(* IEC 61131-3 sources: Lasal-MCP/examples/SampleSource/LASALScreenAdvancedSolution/LASALScreenAdvancedSolution/LASALScreenAdvacnedSolution/Stations/Terminal/HMI/Class/DataRecordSave, 1 file *)

(* ---- DataRecordSave.st ---- *)
(*!
<Class
	Name               = "DataRecordSave"
	Revision           = "0.0"
	RealtimeTask       = "false"
	CyclicTask         = "false"
	BackgroundTask     = "false"
	Sigmatek           = "false"
	OSInterface        = "false"
	HighPriority       = "false"
	Automatic          = "false"
	UpdateMode         = "Prescan"
	SharedCommandTable = "true"
	Objectsize         = "(450,360)">
	<Channels>
		<Server Name="Clear" Visualized="true" Initialize="false" WriteProtected="false" Retentive="false"/>
		<Server Name="IntError" Visualized="false" Initialize="false" WriteProtected="true" Retentive="false"/>
		<Server Name="Load" Visualized="true" Initialize="false" WriteProtected="false" Retentive="false"/>
		<Server Name="Save" Visualized="true" Initialize="false" WriteProtected="false" Retentive="false"/>
		<Server Name="xKoord" Visualized="false" Initialize="false" WriteProtected="true" Retentive="false"/>
		<Server Name="yKoord" Visualized="false" Initialize="false" WriteProtected="true" Retentive="false"/>
		<Client Name="_Grafix" Required="false" Internal="false"/>
		<Client Name="_StdLib" Required="false" Internal="false"/>
		<Client Name="AllocateSize" Required="false" Internal="false" DefValue="4 KB"/>
		<Client Name="FileHandling" Required="true" Internal="false"/>
		<Client Name="FileRead" Required="true" Internal="false"/>
	</Channels>
	<Network Name="DataRecordSave">
		<!-- List of Components in this network -->
		<Components>
			<Object
				Name       = "_base"
				Class      = "_MyIO"
				Position   = "(218,120)"
				Visualized = "true"
				Remotely   = "true">
				<Channels>
					<Server Name="Refresh"/>
					<Server Name="Server0"/>
					<Client Name="Graphic"/>
					<Client Name="Lse"/>
				</Channels>
			</Object>
		</Components>
		<Comments>
		</Comments>
		<!-- List of Connections in this network -->
		<Connections>
			<Connection Source="this.Server0" Destination="_base.Server0" Vertices="(706,210),(534,210),"/>
			<Connection Source="this.Refresh" Destination="_base.Refresh" Vertices="(706,270),(534,270),"/>
			<Connection Source="_base.Lse" Destination="this.Lse" Vertices="(218,210),(38,210),"/>
		</Connections>
		<!-- Headerfiles -->
		<Options>
		</Options>
	</Network>
</Class>
*)
#pragma using _MyIO

DataRecordSave : CLASS
: _MyIO
  //Servers:
	xKoord 	: SvrCh_DINT;
	yKoord 	: SvrCh_DINT;
	IntError 	: SvrCh_DINT;
	Save 	: SvrCh_DINT;
	Load 	: SvrCh_DINT;
	Clear 	: SvrCh_DINT;
  //Clients:
	_Grafix 	: CltChCmd__Grafix;
	_StdLib 	: CltChCmd__StdLib;
	AllocateSize 	: CltCh_UDINT;
	FileRead 	: CltChCmd_FileRead;
	FileHandling 	: CltChCmd_FileHandling;
  //Variables:
		bgColor 	: _COLOR;
		RecordColor 	: _COLOR;
		Del 	: DINT;
		pAct 	: ^_DOT;
		pCheck 	: ^_DOT;
		pNext 	: ^_DOT;
		pStart 	: ^_DOT;
		Buffer 	: UDINT;
		BufferCounter 	: UDINT;
		MaxBufferEntries 	: UDINT;
		pData 	: ^_DOT;
		FileIsRead 	: BOOL;
		Retcode 	: DINT;
		pError 	: ^void;
  //Functions:

	FUNCTION VIRTUAL GLOBAL Init;
				//! <Function Comment="this method will be called once when the focus will be given to this object" Name="GetFocus"/>
	FUNCTION __CDECL VIRTUAL GLOBAL GetFocus
		VAR_INPUT
			pio 	: ^_IO;			//! <Variable Comment="pointer to _IO information" Name="GetFocus.pio"/>
		END_VAR
		VAR_OUTPUT
			retcode (EAX) 	: _DOIT;			//! <Variable Comment="return _IFAILED if you dont want to get the focus on the other hand _IDLE" Name="GetFocus.retcode"/>
		END_VAR;
				//! <Function Comment="this method is called everytime when the input is active and a event occured" Name="GetEvent"/>
	FUNCTION __CDECL VIRTUAL GLOBAL GetEvent
		VAR_INPUT
			ped 	: ^_EDITOR;			//! <Variable Comment="pointer to _EDITOR information" Name="GetEvent.ped"/>
			pe 	: ^_EVENT;			//! <Variable Comment="pointer to _EVENT information" Name="GetEvent.pe"/>
		END_VAR
		VAR_OUTPUT
			retcode (EAX) 	: _DOIT;			//! <Variable Comment="for the returnstatement there are 3 different possibilities&#13;&#10;  _IDLE ..... the system should goon like it is (system goes on)&#13;&#10;  _IDIDIT ... i did it (system is ready)&#13;&#10;  _IFAILED .. i tried to do my best, but i failed (system is ready)&#13;&#10;" Name="GetEvent.retcode"/>
		END_VAR;
				//! <Function Comment="this method is called everytime when system wants to redraw the io" Name="Draw"/>
	FUNCTION __CDECL VIRTUAL GLOBAL Draw
		VAR_INPUT
			pio 	: ^_IO;			//! <Variable Comment="pointer to _IO information" Name="Draw.pio"/>
			pr 	: ^_RESULT;			//! <Variable Comment="pointer to _RESULT information" Name="Draw.pr"/>
			pv 	: ^_VARIABLE;			//! <Variable Comment="pointer to io _VARIABLE information" Name="Draw.pv"/>
			input 	: BOOL;			//! <Variable Comment="TRUE it&apos;s an input&#13;&#10;FALSE it&apos;s an output" Name="Draw.input"/>
		END_VAR
		VAR_OUTPUT
			retcode (EAX) 	: _DOIT;			//! <Variable Comment="for the returnstatement there are 3 different possibilities&#13;&#10;  _IDLE ..... the system should goon like it is (system goes on)&#13;&#10;  _IDIDIT ... i did it (system is ready)&#13;&#10;  _IFAILED .. i tried to do my best, but i failed (system is re" Name="Draw.retcode"/>
		END_VAR;
				//! <Function Comment="this method is called everytime when system wants to get data for defined io.&#13;&#10;&#13;&#10;pr ........ &#13;&#10;pio ....... pointer to io information&#13;&#10;pv ........ pointer to io variableinformation&#13;&#10;input ..... TRUE it&apos;s an input / FALSE it&apos;s an output&#13;&#10;&#13;&#10;for the returnstatement there are 3 different possibilities&#13;&#10;_IDLE ..... the system should goon like it is (system goes on)&#13;&#10;_IDIDIT ... i did it (system is ready)&#13;&#10;_IFAILED .. i tried to do my best, but i failed (system is ready)&#13;&#10;&#13;&#10;if you want to do it let&apos;s return _IDIDIT and initialize the  structure _RESULT&#13;&#10;" Name="GetData"/>
	FUNCTION __CDECL VIRTUAL GLOBAL GetData
		VAR_INPUT
			pr 	: ^_RESULT;			//! <Variable Comment="pointer to _RESULT information" Name="GetData.pr"/>
			pio 	: ^_IO;			//! <Variable Comment="pointer to _IO information" Name="GetData.pio"/>
			pv 	: ^_VARIABLE;			//! <Variable Comment="pointer to _VARIABLE information given by LSE" Name="GetData.pv"/>
			input 	: BOOL;			//! <Variable Comment="TRUE it&apos;s an input&#13;&#10;FALSE it&apos;s an output" Name="GetData.input"/>
		END_VAR
		VAR_OUTPUT
			retcode (EAX) 	: _DOIT;			//! <Variable Comment="for the returnstatement there are 3 different possibilities&#13;&#10;  _IDLE ..... the system should goon like it is (system goes on)&#13;&#10;  _IDIDIT ... i did it (system is ready)&#13;&#10;  _IFAILED .. i tried to do my best, but i failed (system is ready)" Name="GetData.retcode"/>
		END_VAR;
				//! <Function Comment="method is called cyclic during object is on screen&#13;&#10;&#13;&#10;pio ....... &#13;&#10;input .... TRUE it&apos;s an input / FALSE it&apos;s an output&#13;&#10;" Name="IF_Run"/>
	FUNCTION __CDECL VIRTUAL GLOBAL IF_Run
		VAR_INPUT
			pio 	: ^_IO;			//! <Variable Comment="pointer to _IO information given by LSE" Name="IF_Run.pio"/>
			input 	: BOOL;			//! <Variable Comment="TRUE it&apos;s an input&#13;&#10;FALSE it&apos;s an output" Name="IF_Run.input"/>
		END_VAR;

	FUNCTION GLOBAL ClearScreen
		VAR_OUTPUT
			Retcode 	: DINT;
		END_VAR;
  //Tables:
	FUNCTION @STD
		VAR_OUTPUT
			ret_code	: CONFSTATES;
		END_VAR;
	FUNCTION GLOBAL TAB @CT_;
END_CLASS;

#pragma usingLtd _Grafix
#pragma usingLtd _StdLib
#pragma usingLtd FileHandling
#pragma usingLtd FileRead

FUNCTION VIRTUAL GLOBAL DataRecordSave::Init

  if _FirstScan then

    // set buffer to 4KB
    Buffer := AllocateSize;
    MaxBufferEntries := AllocateSize / sizeof(_DOT);

    // allocate memory
    pStart$^void := _StdLib.MallocV1(size0:= Buffer,
                                     mark0:= 0);

    if (pStart = NIL) then
      IntError := -1;
      return;
    else

      pError := _StdLib.MemSet(dest:= pStart,
                               value:= 0,
                               size:= Buffer);

      if (pError <> pStart) then
        IntError := -2;
        return;
      end_if;

    end_if;

    Del := TRUE;
  end_if;

END_FUNCTION

FUNCTION __CDECL VIRTUAL GLOBAL DataRecordSave::GetEvent
	VAR_INPUT
		ped 	: ^_EDITOR;
		pe 	: ^_EVENT;
	END_VAR
	VAR_OUTPUT
		retcode (EAX) 	: _DOIT;
	END_VAR

  _MyIO::GetEvent(ped:=ped, pe:=pe);

  retcode := _IDLE;

  // event hidmove
  if pe^.ftype = _EVENT_HIDMOVE then

    if ((pe^.dot.x > ped^.input.io.space.xy1.x) &
        (pe^.dot.x < ped^.input.io.space.xy2.x) &
        (pe^.dot.y > ped^.input.io.space.xy1.y) &
        (pe^.dot.y < ped^.input.io.space.xy2.y)) then

        Del := FALSE;

        retcode := _IDIDIT;

        // actual coordinates in area
        xKoord := pe^.dot.x - ped^.input.io.space.xy1.x;
        yKoord := pe^.dot.y - ped^.input.io.space.xy1.y;

        // overflow
        if (BufferCounter >= MaxBufferEntries) then
          BufferCounter := 0;

          pAct := pStart;
        end_if;

        pAct^.x := pe^.dot.x;
        pAct^.y := pe^.dot.y;

        pAct := pAct + sizeof(_DOT);
        BufferCounter += 1;

     end_if;

  // event hidrelease
  elsif (pe^.ftype = _EVENT_HIDRELEASE) then
    Del := TRUE;
  end_if;

END_FUNCTION

FUNCTION __CDECL VIRTUAL GLOBAL DataRecordSave::Draw
	VAR_INPUT
		pio 	: ^_IO;
		pr 	: ^_RESULT;
		pv 	: ^_VARIABLE;
		input 	: BOOL;
	END_VAR
	VAR_OUTPUT
		retcode (EAX) 	: _DOIT;
	END_VAR
  VAR
  	act : _NEWSCREEN;
  END_VAR

  _MyIO::Draw(pio:=pio, pr:=pr, pv:=pv, input:=input);

  push_screen(p0:=#act);

  RecordColor := _Grafix.MakeColor(backcolor:= pio^.coltxt,
                                   frontcolor:= pio^.coltxt);

  bgColor := _Grafix.MakeColor(backcolor:= pio^.colback,
                               frontcolor:= pio^.colback);

  // draw background
  if (Del = TRUE) then

      _Grafix.Beam(x0:= pio^.space.xy1.x,
                   y0:= pio^.space.xy1.y,
                   x1:= pio^.space.xy2.x,
                   y1:= pio^.space.xy2.y,
                   attrib:= pio^.attrib,
                   color:= bgColor);
  end_if;

  // place read data on screen
  if FileIsRead = TRUE then

    pStart$^Dint := FileRead.ReadKoords();
    pData := pstart;
    pNext := pData + sizeof(_DOT);

    while ((pData$^Dint <= pStart$^Dint + Buffer) & (FileIsRead = TRUE)) do

      if ((pNext^.x = 0) & (pNext^.y = 0)) then
        pNext := pData;
        FileRead.SetReadState(IsDrawing:=FALSE);
      end_if;

      _Grafix.Line(x0:= pData^.x,
                   y0:= pData^.y,
                   x1:= pNext^.x,
                   y1:= pNext^.y,
                   attrib:= pio^.attrib,
                   color:= RecordColor);

      pData += sizeof(_DOT);
      pNext += sizeof(_dot);

      if (pNext >= pStart + Buffer) then
        pNext := pData;
      end_if;

    end_while;

    FileRead.SetReadState(IsDrawing:= FALSE);

  // draw data on screen
  else

    if (pAct <> NIL) then
      pCheck := pStart;

      while (pCheck < (pAct - sizeof(_DOT))) do

        pNext := pCheck + sizeof(_DOT);

        _Grafix.Line(x0:= pCheck^.x,
                     y0:= pCheck^.y,
                     x1:= pNext^.x,
                     y1:= pNext^.y,
                     attrib:= pio^.attrib,
                     color:= RecordColor);

        pCheck += sizeof(_DOT);

      end_while;

    end_if;
  end_if;

  pop_screen(p0:=#act);
  copy_screen(p0:=#act, p1:=#pio^.space);

  retcode := _IDIDIT;

END_FUNCTION

FUNCTION __CDECL VIRTUAL GLOBAL DataRecordSave::GetFocus
	VAR_INPUT
		pio 	: ^_IO;
	END_VAR
	VAR_OUTPUT
		retcode (EAX) 	: _DOIT;
	END_VAR

  _MyIO::GetFocus(pio:=pio);

  // set pointer to start
  pAct := pStart;
  pCheck  := pStart;
  BufferCounter := 0;

  retcode := _IDLE;

END_FUNCTION

FUNCTION __CDECL VIRTUAL GLOBAL DataRecordSave::IF_Run
	VAR_INPUT
		pio 	: ^_IO;
		input 	: BOOL;
	END_VAR

  _MyIO::IF_Run(pio:=pio, input:=input);

  //****************************************************************
  // save data
  //****************************************************************
  if (Save = 1) then
    Save := 0;
    Retcode := FileHandling.StartWrite(pData:= pStart$^DINT,
                                       Amount:= Buffer);

    if (Retcode < 0) then
      IntError := -2;
      return;
    end_if;

     Refresh := 1;
  end_if;

  //***************************************************************
  // load data
  //***************************************************************
  if (Load = 1) then
    FileRead.StartRead := 1;
    Load := 0;

    if (Retcode < 0) then
      IntError := -3;
      return;
    end_if;

     Refresh := 1;
  end_if;

  FileIsRead := FileRead.GetReadState();

  if (FileIsRead = TRUE) then
    Refresh := 1;
  end_if;

  //***************************************************************
  // clear data
  //***************************************************************
  if (Clear = 1) then

    Retcode := ClearScreen();

    if (Retcode < 0) then
      IntError := -4;
      return;
    end_if;

  end_if;

END_FUNCTION

FUNCTION GLOBAL DataRecordSave::ClearScreen
	VAR_OUTPUT
		Retcode 	: DINT;
	END_VAR

  Retcode := 0;

  // clear screen
  if ((_StdLib.MemSet(dest:=pStart,
                      value:=0,
                      size:=Buffer)) <> pStart) then
    Retcode := -1;
    return;
  end_if;

  Refresh:= 1;

END_FUNCTION

FUNCTION __CDECL VIRTUAL GLOBAL DataRecordSave::GetData
	VAR_INPUT
		pr 	: ^_RESULT;
		pio 	: ^_IO;
		pv 	: ^_VARIABLE;
		input 	: BOOL;
	END_VAR
	VAR_OUTPUT
		retcode (EAX) 	: _DOIT;
	END_VAR

  _MyIO::GetData(pr:=pr, pio:=pio, pv:=pv, input:=input);

  // get X- and Y-Coordinates
  pr^.value := to_dint((to_udint(xKoord) shl 16) xor (to_udint(yKoord)));

  retcode := _IDIDIT;

END_FUNCTION
